FUNCTION_BLOCK my_sequencer EXTENDS TcoCore.TcoSequencer

METHOD PROTECTED Main : BOOL
IF TRUE THEN; END_IF;
END_METHOD

END_FUNCTION_BLOCK

(* stored: Version 1.1.0.1, ProductVersion 3.1.4024.9
   POU my_sequencer: Id {9f9584ee-a192-4ce3-b60b-3cc81b968d12}, SpecialFunc None
   Method Main: Id {c80e0315-425c-484c-97dc-501a0fbb701d} *)
